FUNCTION_BLOCK Dosagem_Alcalinizante (* Dosagem de alcalinizante (800): casca sem logica e sem campo - BO-02, DO-04/05 e LIT-03 so com as tags para o OPC UA - HidrycoLib *)
  (* Standard: 61499-2 *)
  (* Version 1.3, 12/11/2026, Hidryco, Hidryco, 1.3: campo na Remota 1 da Subestacao (A6 %I0.96-104 pelo M262_Substacao): BO/DO com cfgFalhaNA (FALHA = TRUE em falha); LIT_800_03 em 4-20 mA (A12 canal 0); LIGA 800-BO-02 em %Q0.15 (M262_Substacao); LIGA 800-DO-04/05 sai em CNF_DOSADORAS (cmdDO04/05, na mudanca e a cada 5 s) para o Utilities do M262_Nereda, que escreve a word 1 do A8. 1.2: LIT_800_03 como sensor de nivel (cfgNivel, m) para a tela DOSAGEM_ALCALINIZANTE. 1.1: carga no gerador: REQ_GERADOR com geradorHabilitaDO04/DO05 e stsGerador (Subestacao HAB_DO_800_04/05 e stsPlantaNoGerador) para DO_800_04/05 (bloqueio e raio do Motor_Generico). 1.0: casca para a IO List da Nereda (caminhos DosagemAlcalinizante.BO_800_02/DO_800_04/DO_800_05/LIT_800_03). Sem logica e sem campo: motores com cfgUsaTermica = FALSE e sensor com cfgComunicacao = TRUE para nao gerar alarme. Ao ligar o campo, rever esses parametros. *)
  PACKAGE Hidryco.HidrycoLib;
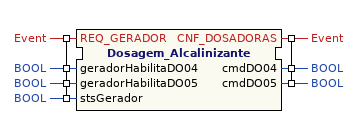
  EVENT_INPUT
    REQ_GERADOR WITH geradorHabilitaDO04, geradorHabilitaDO05, stsGerador; (* Planta no gerador e liberacao das dosadoras (Subestacao) *)
  END_EVENT
  EVENT_OUTPUT
    CNF_DOSADORAS WITH cmdDO04, cmdDO05; (* Comando das dosadoras para o M262_Nereda (Utilities.REQ_DOSADORAS, A8 %Q0.16/17): na mudanca e a cada 5 s *)
  END_EVENT
  VAR_INPUT
    geradorHabilitaDO04 : BOOL; (* 800-DO-04 liberada para operar com a planta nos geradores *)
    geradorHabilitaDO05 : BOOL; (* 800-DO-05 liberada para operar com a planta nos geradores *)
    stsGerador : BOOL; (* TRUE = planta alimentada pelos geradores *)
  END_VAR
  VAR_OUTPUT
    cmdDO04 : BOOL; (* LIGA 800-DO-04 (cmdAcionamento do DO_800_04) *)
    cmdDO05 : BOOL; (* LIGA 800-DO-05 (cmdAcionamento do DO_800_05) *)
  END_VAR
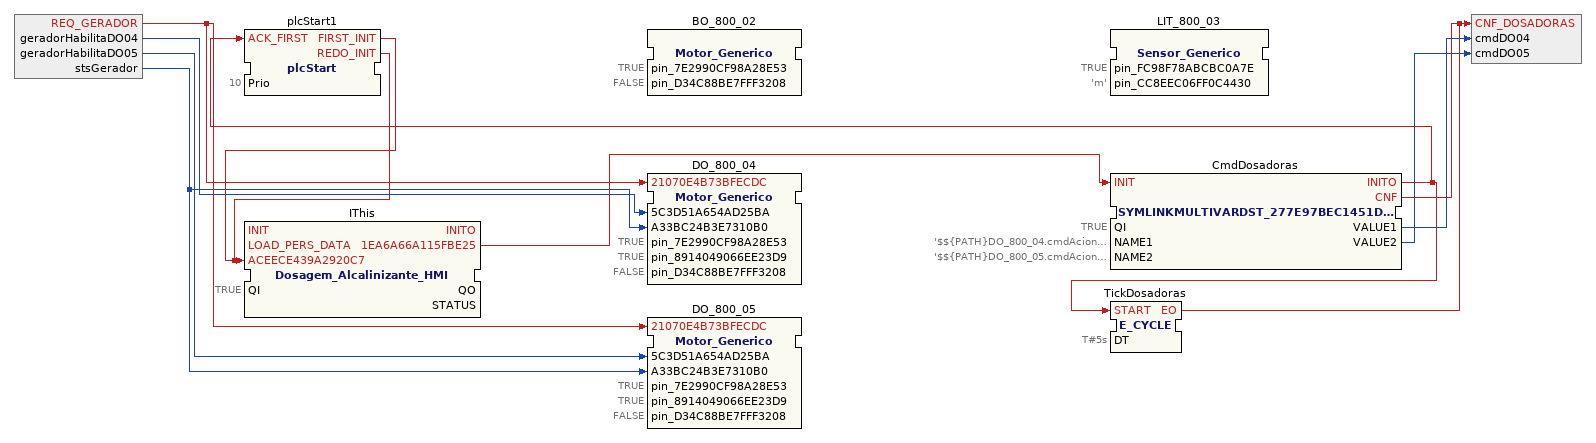
  FBS
    IThis : Dosagem_Alcalinizante_HMI(QI := TRUE);
    plcStart1 : plcStart(Prio := 10);
    BO_800_02 : Motor_Generico(pin_7E2990CF98A28E53 := TRUE, pin_D34C88BE7FFF3208 := FALSE);
    DO_800_04 : Motor_Generico(pin_7E2990CF98A28E53 := TRUE, pin_8914049066EE23D9 := TRUE, pin_D34C88BE7FFF3208 := FALSE);
    DO_800_05 : Motor_Generico(pin_7E2990CF98A28E53 := TRUE, pin_8914049066EE23D9 := TRUE, pin_D34C88BE7FFF3208 := FALSE);
    LIT_800_03 : Sensor_Generico(pin_FC98F78ABCBC0A7E := TRUE, pin_CC8EEC06FF0C4430 := 'm');
    CmdDosadoras : SYMLINKMULTIVARDST_277E97BEC1451D2C(QI := TRUE, NAME1 := '$${PATH}DO_800_04.cmdAcionamento', NAME2 := '$${PATH}DO_800_05.cmdAcionamento'); {SET_ATTRIBUTE(Configuration.GenericFBType.InterfaceParams, Runtime.System#I:=2;VALUE${I$}:BOOL,BOOL)}
    TickDosadoras : E_CYCLE(DT := T#5s);
  END_FBS
  EVENT_CONNECTIONS
    plcStart1.FIRST_INIT TO IThis.ACEECE439A2920C7;
    plcStart1.REDO_INIT TO IThis.ACEECE439A2920C7;
    IThis.1EA6A66A115FBE25 TO CmdDosadoras.INIT;
    CmdDosadoras.INITO TO plcStart1.ACK_FIRST;
    CmdDosadoras.INITO TO TickDosadoras.START;
    CmdDosadoras.CNF TO CNF_DOSADORAS;
    TickDosadoras.EO TO CNF_DOSADORAS;
    REQ_GERADOR TO DO_800_04.21070E4B73BFECDC;
    REQ_GERADOR TO DO_800_05.21070E4B73BFECDC;
  END_CONNECTIONS
  DATA_CONNECTIONS
    geradorHabilitaDO04 TO DO_800_04.5C3D51A654AD25BA;
    geradorHabilitaDO05 TO DO_800_05.5C3D51A654AD25BA;
    stsGerador TO DO_800_04.A33BC24B3E7310B0;
    stsGerador TO DO_800_05.A33BC24B3E7310B0;
    CmdDosadoras.VALUE1 TO cmdDO04;
    CmdDosadoras.VALUE2 TO cmdDO05;
  END_CONNECTIONS
END_FUNCTION_BLOCK
